PROGRAM MAIN
VAR
    fbMotor : FB_Motor;
END_VAR

fbMotor(bEnable := TRUE);

END_PROGRAM

(* stored: Version 1.1.0.1, ProductVersion 3.1.4024.12
   POU MAIN: Id {55555555-0000-0000-0000-000000000001}, SpecialFunc None *)
